(* IEC 61131-3 sources: llm-plc-st-eval/data/definitivo/gpt-4o-2024-08-06/A1/zero_shot, 3 files *)

(* ---- ejec_1.st ---- *)
```pascal
FUNCTION_BLOCK FB_PID
VAR_INPUT
    SP : REAL;      // Setpoint
    PV : REAL;      // Process Variable
    Kp : REAL;      // Proportional Gain
    Ti : REAL;      // Integral Time (seconds)
    Td : REAL;      // Derivative Time (seconds)
    ciclo : TIME;   // Sampling period
END_VAR

VAR_OUTPUT
    CV : REAL;      // Control Variable (output)
END_VAR

VAR
    e : REAL;               // Error
    e_prev : REAL;          // Previous error
    integral : REAL;        // Integral term
    derivative : REAL;      // Derivative term
    dt : REAL;              // Sampling period in seconds
    CV_unsat : REAL;        // Unsaturated control variable
END_VAR

VAR CONSTANT
    CV_MIN : REAL := 0.0;   // Minimum CV
    CV_MAX : REAL := 100.0; // Maximum CV
END_VAR

// Convert TIME to seconds
dt := TO_REAL(ciclo) / 1000.0;

// Calculate error
e := SP - PV;

// Proportional term
CV_unsat := Kp * e;

// Integral term
IF Ti > 0.0 THEN
    integral := integral + (e * dt / Ti);

    // Anti-windup: Clamping
    IF CV_unsat >= CV_MAX THEN
        IF e > 0.0 THEN
            integral := integral - (e * dt / Ti); // Prevent positive windup
        END_IF
    ELSIF CV_unsat <= CV_MIN THEN
        IF e < 0.0 THEN
            integral := integral - (e * dt / Ti); // Prevent negative windup
        END_IF
    END_IF
END_IF

// Add integral term
CV_unsat := CV_unsat + Kp * integral;

// Derivative term
derivative := Td * (e - e_prev) / dt;
CV_unsat := CV_unsat + Kp * derivative;

// Update previous error
e_prev := e;

// Saturate CV
IF CV_unsat > CV_MAX THEN
    CV := CV_MAX;
ELSIF CV_unsat < CV_MIN THEN
    CV := CV_MIN;
ELSE
    CV := CV_unsat;
END_IF

END_FUNCTION_BLOCK
```

(* ---- ejec_2.st ---- *)
```pascal
FUNCTION_BLOCK FB_PID
VAR_INPUT
    SP : REAL;       // Setpoint
    PV : REAL;       // Process Variable
    Kp : REAL;       // Proportional Gain
    Ti : REAL;       // Integral Time (seconds)
    Td : REAL;       // Derivative Time (seconds)
    ciclo : TIME;    // Sampling period
END_VAR

VAR_OUTPUT
    CV : REAL;       // Control Variable (Output)
END_VAR

VAR
    e : REAL;        // Error
    e_prev : REAL;   // Previous error
    integral : REAL; // Integral term
    derivative : REAL; // Derivative term
    dt : REAL;       // Sampling period in seconds
    CV_unsat : REAL; // Unsaturated Control Variable
END_VAR

VAR CONSTANT
    CV_MIN : REAL := 0.0;   // Minimum CV
    CV_MAX : REAL := 100.0; // Maximum CV
END_VAR

// Convert ciclo from TIME to REAL (seconds)
dt := REAL_TO_TIME(ciclo) / 1000.0;

// Calculate error
e := SP - PV;

// Calculate integral term with anti-windup
IF Ti > 0.0 THEN
    integral := integral + e * dt;
    // Anti-windup clamping
    IF CV >= CV_MAX AND e > 0.0 THEN
        integral := integral - e * dt;
    ELSIF CV <= CV_MIN AND e < 0.0 THEN
        integral := integral - e * dt;
    END_IF
ELSE
    integral := 0.0;
END_IF

// Calculate derivative term
derivative := (e - e_prev) / dt;

// Calculate unsaturated CV
CV_unsat := Kp * (e + (1.0 / Ti) * integral + Td * derivative);

// Saturate CV
IF CV_unsat > CV_MAX THEN
    CV := CV_MAX;
ELSIF CV_unsat < CV_MIN THEN
    CV := CV_MIN;
ELSE
    CV := CV_unsat;
END_IF

// Update previous error
e_prev := e;

END_FUNCTION_BLOCK
```

Este código implementa un controlador PID discreto en Structured Text (ST) conforme al estándar IEC 61131-3. El bloque de función `FB_PID` calcula la salida `CV` basada en las entradas proporcionadas, aplicando anti-windup para evitar la acumulación excesiva en el término integral cuando la salida está saturada.

(* ---- ejec_3.st ---- *)
```pascal
FUNCTION_BLOCK FB_PID
VAR_INPUT
    SP : REAL;      // Setpoint
    PV : REAL;      // Process Variable
    Kp : REAL;      // Proportional Gain
    Ti : REAL;      // Integral Time (seconds)
    Td : REAL;      // Derivative Time (seconds)
    ciclo : TIME;   // Sampling Time
END_VAR

VAR_OUTPUT
    CV : REAL;      // Control Variable (0.0 to 100.0)
END_VAR

VAR
    e : REAL;               // Error
    e_prev : REAL;          // Previous Error
    integral : REAL;        // Integral Term
    derivative : REAL;      // Derivative Term
    dt : REAL;              // Sampling Time in seconds
    CV_unsat : REAL;        // Unsaturated Control Variable
END_VAR

VAR CONSTANT
    CV_MIN : REAL := 0.0;   // Minimum CV
    CV_MAX : REAL := 100.0; // Maximum CV
END_VAR

// Convert TIME to seconds
dt := REAL_TO_TIME(ciclo) / 1000.0;

// Calculate error
e := SP - PV;

// Proportional term
CV_unsat := Kp * e;

// Integral term
IF Ti > 0.0 THEN
    integral := integral + (e * dt / Ti);

    // Anti-windup: Clamping
    IF (CV_unsat >= CV_MAX) AND (e > 0.0) THEN
        integral := integral; // Do not accumulate positive error
    ELSIF (CV_unsat <= CV_MIN) AND (e < 0.0) THEN
        integral := integral; // Do not accumulate negative error
    ELSE
        CV_unsat := CV_unsat + Kp * integral;
    END_IF
END_IF

// Derivative term
derivative := Td * (e - e_prev) / dt;
CV_unsat := CV_unsat + Kp * derivative;

// Update previous error
e_prev := e;

// Saturate CV
IF CV_unsat > CV_MAX THEN
    CV := CV_MAX;
ELSIF CV_unsat < CV_MIN THEN
    CV := CV_MIN;
ELSE
    CV := CV_unsat;
END_IF

END_FUNCTION_BLOCK
```

Este código implementa un controlador PID discreto en Structured Text (ST) conforme al estándar IEC 61131-3. El controlador utiliza la forma estándar del PID y aplica técnicas de anti-windup para evitar la acumulación excesiva de la acción integral cuando la salida está saturada.
